// TIA Portal V20 export
Screen "160RobotCollision"  1276x673
  ScreenItem "Graphic view_13" at 333,98 size 634x531  Type=HmiGraphicView
  ScreenItem "矩形_6" at 0,70 size 1274x597  Type=HmiRectangle
  ScreenItem "Graphic view_11" at 331,353 size 410x35  Type=HmiGraphicView
  ScreenItem "Graphic view_12" at 239,353 size 410x35  Type=HmiGraphicView
  ScreenItem "Title_ScreenOverview_X390_Y2" at 438,5 size 551x57  Type=HmiTextBox
  ScreenItem "Line_Header_X0_Y64" at 0,64 size 1274x1  Type=HmiLine
  ScreenItem "permanentareaborderrectangle" at 0,0 size 0x0  Type=HmiRectangle
  ScreenItem "Button_Back" at 2,2 size 90x60  Type=HmiButton
  ScreenItem "Text_5" at 449,616 size 84x39  Type=HmiText
  ScreenItem "Text_6" at 449,77 size 84x39  Type=HmiText
  ScreenItem "Graphic view_6" at 746,-206 size 60x30  Type=HmiGraphicView
  ScreenItem "Graphic view_7" at 746,-594 size 60x30  Type=HmiGraphicView
  ScreenItem "Graphic view_8" at 746,-982 size 60x30  Type=HmiGraphicView
  ScreenItem "Rectangle_6" at 80,259 size 164x328  Type=HmiRectangle
  ScreenItem "Text_75" at 72,257 size 174x35  Type=HmiText
  ScreenItem "Text_76" at 103,283 size 123x35  Type=HmiText
  ScreenItem "Text_77" at 117,311 size 88x35  Type=HmiText
  ScreenItem "Text_78" at 109,339 size 136x35  Type=HmiText
  ScreenItem "矩形_47" at 93,346 size 17x17  Type=HmiRectangle
  ScreenItem "矩形_48" at 93,319 size 17x17  Type=HmiRectangle
  ScreenItem "矩形_49" at 93,292 size 17x17  Type=HmiRectangle
  ScreenItem "Text_83" at 103,393 size 123x35  Type=HmiText
  ScreenItem "Text_84" at 72,367 size 174x35  Type=HmiText
  ScreenItem "矩形_53" at 93,402 size 17x17  Type=HmiRectangle
  ScreenItem "矩形_54" at 93,429 size 17x17  Type=HmiRectangle
  ScreenItem "矩形_55" at 93,456 size 17x17  Type=HmiRectangle
  ScreenItem "Text_85" at 109,449 size 136x35  Type=HmiText
  ScreenItem "Text_86" at 117,421 size 88x35  Type=HmiText
  ScreenItem "Text_1" at 351,209 size 84x60  Type=HmiText
  ScreenItem "Text_2" at 544,461 size 84x60  Type=HmiText
  ScreenItem "Text_3" at 71,473 size 174x35  Type=HmiText
  ScreenItem "矩形_1" at 92,508 size 17x17  Type=HmiRectangle
  ScreenItem "Text_4" at 108,555 size 136x35  Type=HmiText
  ScreenItem "矩形_2" at 92,535 size 17x17  Type=HmiRectangle
  ScreenItem "矩形_3" at 92,562 size 17x17  Type=HmiRectangle
  ScreenItem "Text_7" at 116,527 size 88x35  Type=HmiText
  ScreenItem "Text_8" at 102,499 size 123x35  Type=HmiText
  ScreenItem "Rectangle_1" at 1031,238 size 164x328  Type=HmiRectangle
  ScreenItem "Text_9" at 1023,236 size 174x35  Type=HmiText
  ScreenItem "Text_10" at 1054,262 size 123x35  Type=HmiText
  ScreenItem "Text_11" at 1068,290 size 88x35  Type=HmiText
  ScreenItem "Text_12" at 1060,318 size 136x35  Type=HmiText
  ScreenItem "矩形_4" at 1044,325 size 17x17  Type=HmiRectangle
  ScreenItem "矩形_5" at 1044,298 size 17x17  Type=HmiRectangle
  ScreenItem "矩形_7" at 1044,271 size 17x17  Type=HmiRectangle
  ScreenItem "Text_13" at 1054,372 size 123x35  Type=HmiText
  ScreenItem "Text_14" at 1023,346 size 174x35  Type=HmiText
  ScreenItem "矩形_8" at 1044,381 size 17x17  Type=HmiRectangle
  ScreenItem "矩形_9" at 1044,408 size 17x17  Type=HmiRectangle
  ScreenItem "矩形_10" at 1044,435 size 17x17  Type=HmiRectangle
  ScreenItem "Text_15" at 1060,428 size 136x35  Type=HmiText
  ScreenItem "Text_16" at 1068,400 size 88x35  Type=HmiText
  ScreenItem "Text_17" at 1022,452 size 174x35  Type=HmiText
  ScreenItem "矩形_11" at 1043,487 size 17x17  Type=HmiRectangle
  ScreenItem "Text_18" at 1059,534 size 136x35  Type=HmiText
  ScreenItem "矩形_12" at 1043,514 size 17x17  Type=HmiRectangle
  ScreenItem "矩形_13" at 1043,541 size 17x17  Type=HmiRectangle
  ScreenItem "Text_19" at 1067,506 size 88x35  Type=HmiText
  ScreenItem "Text_20" at 1053,478 size 123x35  Type=HmiText
